(*
SPDX-FileCopyrightText: © 2026 Oleksandr Tiutyk <trofimich@gmail.com>
SPDX-License-Identifier: MIT
License: https://opensource.org/license/mit
*)
(*!
<summary>Identifies owned log discovery, byte readback, deletion and final directory cleanup.</summary>
*)
{attribute 'qualified_only'}
{attribute 'strict'}
TYPE LOGGER_DIRECTORY_CLEANUP_PHASE :
(
	ENUMERATE_FIRST,
	ENUMERATE_WAIT,
	ENUMERATE_NEXT,
	LOAD_FILE,
	WAIT_FOR_LOAD,
	DELETE_FILE,
	WAIT_FOR_DELETE,
	REMOVE_DIRECTORY,
	COMPLETE
);
END_TYPE

(* stored: Version 1.1.0.1
   DUT LOGGER_DIRECTORY_CLEANUP_PHASE: Id {81d3c844-8f9a-407e-86c6-3348aa811116} *)
